Staubli VAL3: CheckTraj.pgx

program CheckTraj(point x_pStart, trsf x_trOffset, point x_pEnd, string x_sMethod, bool& x_bTrajOK)
  local bool l_bOk
  local bool l_bOut
  local num l_nStep
  local trsf l_trMiniOffset
  local trsf l_trStepOffset
  local num l_nVal
  local point l_pTarget
  local jointRx l_jNearBy
  local jointRx l_jTarget
  local jointRx l_jStart
  local point l_pNearBy
  local string l_sPopMsg
begin
  l_trMiniOffset={x_trOffset.x/1000,x_trOffset.y/1000,x_trOffset.z/1000,x_trOffset.rx/1000,x_trOffset.ry/1000,x_trOffset.rz/1000}

  switch x_sMethod
    case "Appro"
      x_pEnd=appro(x_pStart,x_trOffset)
    break
    case "Compose"
      x_pEnd=compose(x_pStart,world,x_trOffset)
      x_pEnd.trsf.x=x_pStart.trsf.x
      x_pEnd.trsf.y=x_pStart.trsf.y
      x_pEnd.trsf.z=x_pStart.trsf.z
    break
  endSwitch


  l_nStep=0
  l_nVal=1
  do
    switch l_nStep
      //******************************************************************
      //Check NearBy Position
      case 0
        l_bOk=pointToJoint(utCurrentTool.tValue,herej(),x_pStart,l_jStart)
        if l_bOk==true
          l_nStep=1
        else
          l_nStep=99
        endIf
      break
      //
      case 1
        switch x_sMethod
          case "Appro"
            l_pNearBy=appro(x_pStart,l_trMiniOffset)
          break
          case "Compose"
            l_pNearBy=compose(x_pStart,world,l_trMiniOffset)
            l_pNearBy.trsf.x=x_pStart.trsf.x
            l_pNearBy.trsf.y=x_pStart.trsf.y
            l_pNearBy.trsf.z=x_pStart.trsf.z
          break
        endSwitch
        l_bOk=pointToJoint(utCurrentTool.tValue,herej(),l_pNearBy,l_jNearBy)
        if l_bOk==true
          l_nStep=2
        else
          l_nStep=99
        endIf
      break
      //******************************************************************
      case 2
        l_trStepOffset={x_trOffset.x*l_nVal/100,x_trOffset.y*l_nVal/100,x_trOffset.z*l_nVal/100,x_trOffset.rx*l_nVal/100,x_trOffset.ry*l_nVal/100,x_trOffset.rz*l_nVal/100}
        switch x_sMethod
          case "Appro"
            l_pTarget=appro(x_pStart,l_trStepOffset)
          break
          case "Compose"
            l_pTarget=compose(x_pStart,world,l_trStepOffset)
            l_pTarget.trsf.x=x_pStart.trsf.x
            l_pTarget.trsf.y=x_pStart.trsf.y
            l_pTarget.trsf.z=x_pStart.trsf.z
          break
        endSwitch
        l_bOk=pointToJoint(utCurrentTool.tValue,herej(),l_pTarget,l_jTarget)
        if l_bOk==true
          l_nStep=3
        else
          l_nStep=99
        endIf
      break
      //
      case 3
        if l_jNearBy.j4-l_jStart.j4>=0 and l_jTarget.j4-l_jStart.j4<0
          l_jTarget.j4=l_jTarget.j4+360
        endIf
        if l_jNearBy.j4-l_jStart.j4<0 and l_jTarget.j4-l_jStart.j4>=0
          l_jTarget.j4=l_jTarget.j4-360
        endIf
        //
        //
        if l_jNearBy.j6-l_jStart.j6>=0 and l_jTarget.j6-l_jStart.j6<0
          l_jTarget.j6=l_jTarget.j6+360
        endIf
        if l_jNearBy.j6-l_jStart.j6<0 and l_jTarget.j6-l_jStart.j6>=0
          l_jTarget.j6=l_jTarget.j6-360
        endIf
        l_nStep=4
      break
      //
      case 4
        if isInRange(l_jTarget)==true
          l_nStep=5
        else
          l_nStep=99
        endIf
      break
      //
      case 5
        if l_nVal<100
          l_nVal=l_nVal+1
          l_nStep=2
        else
          l_nStep=100
        endIf
      break
      //******************************************************************
      case 99
        call updateStr(121,l_sPopMsg,"The maximum rotation angle is only:")
        l_nVal=l_nVal-1
        l_sPopMsg=l_sPopMsg+toString(".",roundDown(l_nVal))+"°"
        popUpMsg(l_sPopMsg)
        //
        x_bTrajOK=false
        l_bOut=true
      break
      case 100
        x_bTrajOK=true
        l_bOut=true
      break
    endSwitch
  until l_bOut
end
